(* IEC 61131-3 sources: plcassist-cli/packages/volt-lsp-iec/test-corpus/lenze-mid/Device/Plc Logic/Application/Library Manager/L_MC1P_MotionControlBasic (part 8) *)

(* ---- MC_READBOOLPARAMETER.fb ---- *)
FUNCTION_BLOCK MC_READBOOLPARAMETER EXTENDS L_MC1P_Template_NoAxis
VAR_INPUT
	AXIS : L_MC1P_IMCParameterAccess;
	ENABLE : BOOL;
	PARAMETERNUMBER : DINT;
END_VAR
VAR_OUTPUT
	VALID : BOOL;
	BUSY : BOOL;
	ERROR : BOOL;
	ERRORID : L_IE1P_Error;
	VALUE : BOOL;
END_VAR
VAR
	XENABLEOLD : BOOL := FALSE;
	PARAMETERNUMBEROLD : DINT := 0;
	L_DCO_READDRIVEPARAMETER1 : L_DCO_ReadDriveParameter;
	TIMERREADCYCLE : TON;
	TCYCLETIME : TIME := TIME#1ms;
	XERRORHOLD : BOOL;
	EERRORIDHOLD : L_IE1P_Error;
	PAXISREF : POINTER TO AXIS_REF;
	PINSTANCE : POINTER TO BYTE;
	EAXISTYPE : L_MC1P_AxisType;
	AXISOLD : L_MC1P_IMCParameterAccess;
	_MCCALL : L_UM1P_MCMultipleCall;
	INPUTDATA : ARRAY [1.._MCCall.c_BufferDepthInput] OF L_MC1P_ReadBoolParameterInput;
	OUTPUTDATA : ARRAY [1.._MCCall.c_BufferDepthOutput] OF L_MC1P_ReadBoolParameterOutput;
	POUTPUTDATA : POINTER TO L_MC1P_ReadBoolParameterOutput;
	XAXISTASKIDXVALID : BOOL;
	ITFSETPOINTINFO : L_UM1P_ISetpointInfo;
	IAXISTASKIDX : INT;
	READCYCLE : TIME;
END_VAR
END_FUNCTION_BLOCK

METHOD FB_RESET : BOOL
END_METHOD

METHOD CALLFUNCTION
VAR_INPUT
	UIINPUTDATAIDX : UINT;
	UIOUTPUTDATAIDX : UINT;
END_VAR
END_METHOD

METHOD COPYINPUTS : BOOL
VAR_INPUT
	IDX : WORD;
END_VAR
END_METHOD

METHOD COPYOUTPUTS : BOOL
VAR_INPUT
	IDX : WORD;
END_VAR
END_METHOD

METHOD FUNCTIONWASCALLEDTWICE : BOOL
VAR_INPUT
	IDX : WORD;
END_VAR
END_METHOD

METHOD HANDLESTANDARDCALL : BOOL
END_METHOD

METHOD SYNCOUTPUTS
VAR_INPUT
	UICOPYOUTPUTFROMIDX : UINT;
	UICOPYOUTPUTTOIDX : UINT;
END_VAR
END_METHOD

(* ---- MC_READMOTIONSTATE.fb ---- *)
FUNCTION_BLOCK MC_READMOTIONSTATE EXTENDS L_MC1P_Template
VAR_INPUT
	ENABLE : BOOL;
	SOURCE : MC_SOURCE;
END_VAR
VAR_OUTPUT
	VALID : BOOL;
	BUSY : BOOL;
	ERROR : BOOL;
	ERRORID : L_IE1P_Error;
	CONSTANTVELOCITY : BOOL;
	ACCELERATING : BOOL;
	DECELERATING : BOOL;
	DIRECTIONPOSITIVE : BOOL;
	DIRECTIONNEGATIVE : BOOL;
	INPOSITION : BOOL;
	STANDSTILLSETVELOCITY : BOOL;
	STANDSTILLACTVELOCITY : BOOL;
END_VAR
VAR
	READ : L_MC1P_ReadMotionState_Internal;
	_MCCALL : L_UM1P_MCMultipleCall;
	INPUTDATA : ARRAY [1.._MCCall.c_BufferDepthInput] OF L_MC1P_ReadMotionStateInput;
	OUTPUTDATA : ARRAY [1.._MCCall.c_BufferDepthOutput] OF L_MC1P_ReadMotionStateOutput;
END_VAR
END_FUNCTION_BLOCK

METHOD CALLFUNCTION
VAR_INPUT
	UIINPUTDATAIDX : UINT;
	UIOUTPUTDATAIDX : UINT;
END_VAR
END_METHOD

METHOD COPYINPUTS : BOOL
VAR_INPUT
	IDX : WORD;
END_VAR
END_METHOD

METHOD COPYOUTPUTS : BOOL
VAR_INPUT
	IDX : WORD;
END_VAR
END_METHOD

METHOD FUNCTIONWASCALLEDTWICE : BOOL
VAR_INPUT
	IDX : WORD;
END_VAR
END_METHOD

METHOD HANDLESTANDARDCALL : BOOL
END_METHOD

METHOD SYNCOUTPUTS
VAR_INPUT
	UICOPYOUTPUTFROMIDX : UINT;
	UICOPYOUTPUTTOIDX : UINT;
END_VAR
END_METHOD

(* ---- MC_READPARAMETER.fb ---- *)
FUNCTION_BLOCK MC_READPARAMETER EXTENDS L_MC1P_Template_NoAxis
VAR_INPUT
	AXIS : L_MC1P_IMCParameterAccess;
	ENABLE : BOOL;
	PARAMETERNUMBER : DINT;
END_VAR
VAR_OUTPUT
	VALID : BOOL;
	BUSY : BOOL;
	ERROR : BOOL;
	ERRORID : L_IE1P_Error;
	VALUE : LREAL;
END_VAR
VAR
	READ : L_MC1P_ReadParameter_Internal;
	TCYCLETIME : TIME := TIME#1ms;
	_MCCALL : L_UM1P_MCMultipleCall;
	INPUTDATA : ARRAY [1.._MCCall.c_BufferDepthInput] OF L_MC1P_ReadParameterInput;
	OUTPUTDATA : ARRAY [1.._MCCall.c_BufferDepthOutput] OF L_MC1P_ReadParameterOutput;
	PINPUTDATA : POINTER TO L_MC1P_ReadParameterInput;
	ITFSETPOINTINFO : L_UM1P_ISetpointInfo;
	XAXISTASKIDXVALID : BOOL;
	IAXISTASKIDX : INT;
	READCYCLE : TIME;
END_VAR
END_FUNCTION_BLOCK

METHOD CALLFUNCTION
VAR_INPUT
	UIINPUTDATAIDX : UINT;
	UIOUTPUTDATAIDX : UINT;
END_VAR
END_METHOD

METHOD COPYINPUTS : BOOL
VAR_INPUT
	IDX : WORD;
END_VAR
END_METHOD

METHOD COPYOUTPUTS : BOOL
VAR_INPUT
	IDX : WORD;
END_VAR
END_METHOD

METHOD FUNCTIONWASCALLEDTWICE : BOOL
VAR_INPUT
	IDX : WORD;
END_VAR
END_METHOD

METHOD HANDLESTANDARDCALL : BOOL
END_METHOD

METHOD SYNCOUTPUTS
VAR_INPUT
	UICOPYOUTPUTFROMIDX : UINT;
	UICOPYOUTPUTTOIDX : UINT;
END_VAR
END_METHOD

(* ---- MC_READSTATUS.fb ---- *)
FUNCTION_BLOCK MC_READSTATUS EXTENDS L_MC1P_Template
VAR_INPUT
	ENABLE : BOOL;
END_VAR
VAR_OUTPUT
	VALID : BOOL;
	BUSY : BOOL;
	ERROR : BOOL;
	ERRORID : L_IE1P_Error;
	ERRORSTOP : BOOL;
	DISABLED : BOOL;
	STOPPING : BOOL;
	HOMING : BOOL;
	STANDSTILL : BOOL;
	DISCRETEMOTION : BOOL;
	CONTINUOUSMOTION : BOOL;
	SYNCHRONIZEDMOTION : BOOL;
	CONSTANTVELOCITY : BOOL;
	ACCELERATING : BOOL;
	DECELERATING : BOOL;
	INPOSITION : BOOL;
END_VAR
VAR
	XENABLEOLD : BOOL := FALSE;
	_MCCALL : L_UM1P_MCMultipleCall;
	INPUTDATA : ARRAY [1.._MCCall.c_BufferDepthInput] OF L_MC1P_ReadStatusInput;
	OUTPUTDATA : ARRAY [1.._MCCall.c_BufferDepthOutput] OF L_MC1P_ReadStatusOutput;
	POUTPUTDATA : POINTER TO L_MC1P_ReadStatusOutput;
END_VAR
END_FUNCTION_BLOCK

METHOD FB_RESET : BOOL
END_METHOD

METHOD CALLFUNCTION
VAR_INPUT
	UIINPUTDATAIDX : UINT;
	UIOUTPUTDATAIDX : UINT;
END_VAR
END_METHOD

METHOD COPYINPUTS : BOOL
VAR_INPUT
	IDX : WORD;
END_VAR
END_METHOD

METHOD COPYOUTPUTS : BOOL
VAR_INPUT
	IDX : WORD;
END_VAR
END_METHOD

METHOD FUNCTIONWASCALLEDTWICE : BOOL
VAR_INPUT
	IDX : WORD;
END_VAR
END_METHOD

METHOD HANDLESTANDARDCALL : BOOL
END_METHOD

METHOD SYNCOUTPUTS
VAR_INPUT
	UICOPYOUTPUTFROMIDX : UINT;
	UICOPYOUTPUTTOIDX : UINT;
END_VAR
END_METHOD

(* ---- MC_RESET.fb ---- *)
FUNCTION_BLOCK MC_RESET EXTENDS L_MC1P_Template
VAR_INPUT
	EXECUTE : BOOL;
END_VAR
VAR_OUTPUT
	DONE : BOOL;
	BUSY : BOOL;
	ERROR : BOOL;
	ERRORID : L_IE1P_Error;
END_VAR
VAR
	RESET : L_MC1P_Reset_Internal;
	RESETINPUT : L_MC1P_ResetInput;
	RESETOUTPUT : L_MC1P_ResetOutput;
	_MCCALL : L_UM1P_MCMultipleCall := STRUCT(itfMCCall := THIS^);
	INPUTDATA : ARRAY [1.._MCCall.c_BufferDepthInput] OF L_MC1P_ResetInput;
	OUTPUTDATA : ARRAY [1.._MCCall.c_BufferDepthOutput] OF L_MC1P_ResetOutput;
	POUTPUTDATA : POINTER TO L_MC1P_ResetOutput;
END_VAR
END_FUNCTION_BLOCK

METHOD CALLFUNCTION
VAR_INPUT
	UIINPUTDATAIDX : UINT;
	UIOUTPUTDATAIDX : UINT;
END_VAR
END_METHOD

METHOD COPYINPUTS : BOOL
VAR_INPUT
	IDX : WORD;
END_VAR
END_METHOD

METHOD COPYOUTPUTS : BOOL
VAR_INPUT
	IDX : WORD;
END_VAR
END_METHOD

METHOD FUNCTIONWASCALLEDTWICE : BOOL
VAR_INPUT
	IDX : WORD;
END_VAR
END_METHOD

METHOD HANDLESTANDARDCALL : BOOL
END_METHOD

METHOD SYNCOUTPUTS
VAR_INPUT
	UICOPYOUTPUTFROMIDX : UINT;
	UICOPYOUTPUTTOIDX : UINT;
END_VAR
END_METHOD

(* ---- MC_SETOVERRIDE.fb ---- *)
FUNCTION_BLOCK MC_SETOVERRIDE EXTENDS L_MC1P_Template
VAR_INPUT
	ENABLE : BOOL;
	VELFACTOR : LREAL := 1.0;
	ACCFACTOR : LREAL := 1.0;
	JERKFACTOR : LREAL := 1.0;
END_VAR
VAR_OUTPUT
	ENABLED : BOOL;
	BUSY : BOOL;
	ERROR : BOOL;
	ERRORID : L_IE1P_Error;
END_VAR
VAR
	OVERRIDE : L_MC1P_SetOverride_Internal;
	_MCCALL : L_UM1P_MCMultipleCall;
	INPUTDATA : ARRAY [1.._MCCall.c_BufferDepthInput] OF L_MC1P_SetOverrideInput;
	OUTPUTDATA : ARRAY [1.._MCCall.c_BufferDepthOutput] OF L_MC1P_SetOverrideOutput;
END_VAR
END_FUNCTION_BLOCK

METHOD CALLFUNCTION
VAR_INPUT
	UIINPUTDATAIDX : UINT;
	UIOUTPUTDATAIDX : UINT;
END_VAR
END_METHOD

METHOD COPYINPUTS : BOOL
VAR_INPUT
	IDX : WORD;
END_VAR
END_METHOD

METHOD COPYOUTPUTS : BOOL
VAR_INPUT
	IDX : WORD;
END_VAR
END_METHOD

METHOD FUNCTIONWASCALLEDTWICE : BOOL
VAR_INPUT
	IDX : WORD;
END_VAR
END_METHOD

METHOD HANDLESTANDARDCALL : BOOL
END_METHOD

METHOD SYNCOUTPUTS
VAR_INPUT
	UICOPYOUTPUTFROMIDX : UINT;
	UICOPYOUTPUTTOIDX : UINT;
END_VAR
END_METHOD

(* ---- MC_SETPOSITION.fb ---- *)
FUNCTION_BLOCK MC_SETPOSITION EXTENDS L_MC1P_Template
VAR_INPUT
	EXECUTE : BOOL;
	POSITION : LREAL;
	RELATIVE : BOOL;
	EXECUTIONMODE : MC_EXECUTION_MODE := MC_EXECUTION_MODE.mcImmediately;
	RESTARTPOSITIONING : BOOL := FALSE;
	USESETTINGSFROMHOMINGMODE : BOOL := FALSE;
END_VAR
VAR_OUTPUT
	DONE : BOOL;
	BUSY : BOOL;
	ERROR : BOOL;
	ERRORID : L_IE1P_Error;
END_VAR
VAR
	XEXECUTEOLD : BOOL;
	XCALLFROMAXESGROUP : BOOL;
	LRDUMMY : LREAL;
	XDISABLELOGMESSAGE : BOOL := FALSE;
	_MCCALL : L_UM1P_MCMultipleCall;
	INPUTDATA : ARRAY [1.._MCCall.c_BufferDepthInput] OF L_MC1P_SetPositionInput;
	OUTPUTDATA : ARRAY [1.._MCCall.c_BufferDepthOutput] OF L_MC1P_SetPositionOutput;
	DISABLELOGMESSAGE : BOOL;
END_VAR
END_FUNCTION_BLOCK

METHOD SETCALLFROMAXESGROUP
VAR_INPUT
	XSETCALLFROMAXESGROUP : BOOL;
END_VAR
END_METHOD

METHOD CALLFUNCTION
VAR_INPUT
	UIINPUTDATAIDX : UINT;
	UIOUTPUTDATAIDX : UINT;
END_VAR
END_METHOD

METHOD COPYINPUTS : BOOL
VAR_INPUT
	IDX : WORD;
END_VAR
END_METHOD

METHOD COPYOUTPUTS : BOOL
VAR_INPUT
	IDX : WORD;
END_VAR
END_METHOD

METHOD FUNCTIONWASCALLEDTWICE : BOOL
VAR_INPUT
	IDX : WORD;
END_VAR
END_METHOD

METHOD HANDLESTANDARDCALL : BOOL
END_METHOD

METHOD SYNCOUTPUTS
VAR_INPUT
	UICOPYOUTPUTFROMIDX : UINT;
	UICOPYOUTPUTTOIDX : UINT;
END_VAR
END_METHOD

(* ---- MC_STOP.fb ---- *)
FUNCTION_BLOCK MC_STOP EXTENDS L_MC1P_Template_Licence_150
VAR_INPUT
	EXECUTE : BOOL;
	DECELERATION : LREAL;
	JERK : LREAL;
END_VAR
VAR_OUTPUT
	DONE : BOOL;
	BUSY : BOOL;
	COMMANDABORTED : BOOL;
	ERROR : BOOL;
	ERRORID : L_IE1P_Error;
END_VAR
VAR
	STOP : L_MC1P_Stop_Internal;
	_MCCALL : L_UM1P_MCMultipleCall;
	INPUTDATA : ARRAY [1.._MCCall.c_BufferDepthInput] OF L_MC1P_StopInput;
	OUTPUTDATA : ARRAY [1.._MCCall.c_BufferDepthOutput] OF L_MC1P_StopOutput;
	PROFILETIME : TIME;
	REMAININGTIMEOFPROFILE : LREAL;
	REMAININGTIMEOFPROFILEAVAILABLE : BOOL;
END_VAR
END_FUNCTION_BLOCK

METHOD CALLFUNCTION
VAR_INPUT
	UIINPUTDATAIDX : UINT;
	UIOUTPUTDATAIDX : UINT;
END_VAR
END_METHOD

METHOD COPYINPUTS : BOOL
VAR_INPUT
	IDX : WORD;
END_VAR
END_METHOD

METHOD COPYOUTPUTS : BOOL
VAR_INPUT
	IDX : WORD;
END_VAR
END_METHOD

METHOD FUNCTIONWASCALLEDTWICE : BOOL
VAR_INPUT
	IDX : WORD;
END_VAR
END_METHOD

METHOD HANDLESTANDARDCALL : BOOL
END_METHOD

METHOD SYNCOUTPUTS
VAR_INPUT
	UICOPYOUTPUTFROMIDX : UINT;
	UICOPYOUTPUTTOIDX : UINT;
END_VAR
END_METHOD

(* ---- MC_TOUCHPROBE.fb ---- *)
FUNCTION_BLOCK MC_TOUCHPROBE EXTENDS L_MC1P_Template
VAR_INPUT
	EXECUTE : BOOL;
	WINDOWONLY : BOOL;
	FIRSTPOSITION : LREAL;
	LASTPOSITION : LREAL;
END_VAR
VAR_OUTPUT
	DONE : BOOL;
	BUSY : BOOL;
	COMMANDABORTED : BOOL;
	ERROR : BOOL;
	ERRORID : L_IE1P_Error;
	ACTIVATIONLEVEL : BOOL;
	ACTIVATIONLEVELVALID : BOOL;
	VALUESTORED_POSEDGE : BOOL;
	RECPOSITION_POSEDGE : LREAL;
	VALUESTORED_NEGEDGE : BOOL;
	RECPOSITION_NEGEDGE : LREAL;
	NEWVALUESTORED_POSEDGE : BOOL;
	NEWVALUESTORED_NEGEDGE : BOOL;
	RECDATA : L_MC1P_TpReceiveData;
END_VAR
VAR_IN_OUT
	TRIGGERINPUT : MC_TRIGGER_REF;
END_VAR
VAR
	TP : L_MC1P_TouchProbe_Internal;
	_MCCALL : L_UM1P_MCMultipleCall := STRUCT(itfMCCall := THIS^);
	INPUTDATA : ARRAY [1.._MCCall.c_BufferDepthInput] OF L_MC1P_TouchProbeInput;
	OUTPUTDATA : ARRAY [1.._MCCall.c_BufferDepthOutput] OF L_MC1P_TouchProbeOutput;
	_FB_SEMA : L_MC1P_CriticalSection;
	_DWUPDATETIME : DWORD;
	DWACTTIMESTAMPSAVE : DWORD;
	XMULTICOREOPTION : BOOL;
END_VAR
END_FUNCTION_BLOCK

METHOD GETACTTPRECEIVEDATA : L_MC1P_TpReceiveData
END_METHOD

METHOD ISUPTODATE : BOOL
VAR_INPUT
	DWUPDATETIME : DWORD;
END_VAR
END_METHOD

METHOD RECDATAISVALID : BOOL
VAR_IN_OUT
	SCRECDATA : L_MC1P_TpReceiveData;
END_VAR
END_METHOD

METHOD REQUESTINTERFACE : BOOL
VAR_INPUT
	ID : DINT;
	PITFUNKNOWN : POINTER TO L_UBUP_IUnknown;
END_VAR
END_METHOD

METHOD CALLFUNCTION
VAR_INPUT
	UIINPUTDATAIDX : UINT;
	UIOUTPUTDATAIDX : UINT;
END_VAR
END_METHOD

METHOD COPYINPUTS : BOOL
VAR_INPUT
	IDX : WORD;
END_VAR
END_METHOD

METHOD COPYOUTPUTS : BOOL
VAR_INPUT
	IDX : WORD;
END_VAR
END_METHOD

METHOD FUNCTIONWASCALLEDTWICE : BOOL
VAR_INPUT
	IDX : WORD;
END_VAR
END_METHOD

METHOD HANDLESTANDARDCALL : BOOL
END_METHOD

METHOD SYNCOUTPUTS
VAR_INPUT
	UICOPYOUTPUTFROMIDX : UINT;
	UICOPYOUTPUTTOIDX : UINT;
END_VAR
END_METHOD

(* ---- MC_WRITEBOOLPARAMETER.fb ---- *)
FUNCTION_BLOCK MC_WRITEBOOLPARAMETER EXTENDS L_MC1P_Template_NoAxis
VAR_INPUT
	AXIS : L_MC1P_IMCParameterAccess;
	EXECUTE : BOOL;
	PARAMETERNUMBER : DINT;
	VALUE : BOOL;
	EXECUTIONMODE : MC_EXECUTION_MODE;
END_VAR
VAR_OUTPUT
	DONE : BOOL;
	BUSY : BOOL;
	ERROR : BOOL;
	ERRORID : L_IE1P_Error;
END_VAR
VAR
	XEXECUTEOLD : BOOL := FALSE;
	XRESETOUTPUT : BOOL := FALSE;
	L_DCO_WRITEDRIVEPARAMETER1 : L_DCO_WriteDriveParameter;
	WERRORID_INT : WORD;
	AXISOLD : L_MC1P_IMCParameterAccess;
	PAXISREF : POINTER TO AXIS_REF;
	XWRITEPARAMETER : BOOL;
	PINSTANCE : POINTER TO BYTE;
	EAXISTYPE : L_MC1P_AxisType;
	_MCCALL : L_UM1P_MCMultipleCall;
	INPUTDATA : ARRAY [1.._MCCall.c_BufferDepthInput] OF L_MC1P_WriteBoolParameterInput;
	OUTPUTDATA : ARRAY [1.._MCCall.c_BufferDepthOutput] OF L_MC1P_WriteBoolParameterOutput;
	POUTPUTDATA : POINTER TO L_MC1P_WriteBoolParameterOutput;
	ITFSETPOINTINFO : L_UM1P_ISetpointInfo;
	XAXISTASKIDXVALID : BOOL;
	IAXISTASKIDX : INT;
END_VAR
END_FUNCTION_BLOCK

METHOD FB_RESET : BOOL
END_METHOD

METHOD CALLFUNCTION
VAR_INPUT
	UIINPUTDATAIDX : UINT;
	UIOUTPUTDATAIDX : UINT;
END_VAR
END_METHOD

METHOD COPYINPUTS : BOOL
VAR_INPUT
	IDX : WORD;
END_VAR
END_METHOD

METHOD COPYOUTPUTS : BOOL
VAR_INPUT
	IDX : WORD;
END_VAR
END_METHOD

METHOD FUNCTIONWASCALLEDTWICE : BOOL
VAR_INPUT
	IDX : WORD;
END_VAR
END_METHOD

METHOD HANDLESTANDARDCALL : BOOL
END_METHOD

METHOD SYNCOUTPUTS
VAR_INPUT
	UICOPYOUTPUTFROMIDX : UINT;
	UICOPYOUTPUTTOIDX : UINT;
END_VAR
END_METHOD

(* ---- MC_WRITEPARAMETER.fb ---- *)
FUNCTION_BLOCK MC_WRITEPARAMETER EXTENDS L_MC1P_Template_NoAxis
VAR_INPUT
	AXIS : L_MC1P_IMCParameterAccess;
	EXECUTE : BOOL;
	PARAMETERNUMBER : DINT;
	VALUE : LREAL;
	EXECUTIONMODE : MC_EXECUTION_MODE;
END_VAR
VAR_OUTPUT
	DONE : BOOL;
	BUSY : BOOL;
	ERROR : BOOL;
	ERRORID : L_IE1P_Error;
END_VAR
VAR
	XEXECUTEOLD : BOOL := FALSE;
	XRESETOUTPUT : BOOL := FALSE;
	AXISOLD : L_MC1P_IMCParameterAccess;
	L_DCO_WRITEDRIVEPARAMETER1 : L_DCO_WriteDriveParameter;
	DWPARAMETERNUMBERINT : DWORD;
	WERRORID_INT : WORD;
	PAXISREF : POINTER TO AXIS_REF;
	PINSTANCE : POINTER TO BYTE;
	EAXISTYPE : L_MC1P_AxisType;
	_MCCALL : L_UM1P_MCMultipleCall;
	INPUTDATA : ARRAY [1.._MCCall.c_BufferDepthInput] OF L_MC1P_WriteParameterInput;
	OUTPUTDATA : ARRAY [1.._MCCall.c_BufferDepthOutput] OF L_MC1P_WriteParameterOutput;
	POUTPUTDATA : POINTER TO L_MC1P_WriteParameterOutput;
	ITFSETPOINTINFO : L_UM1P_ISetpointInfo;
	XAXISTASKIDXVALID : BOOL;
	IAXISTASKIDX : INT;
END_VAR
END_FUNCTION_BLOCK

METHOD FB_RESET : BOOL
END_METHOD

METHOD CALLFUNCTION
VAR_INPUT
	UIINPUTDATAIDX : UINT;
	UIOUTPUTDATAIDX : UINT;
END_VAR
END_METHOD

METHOD COPYINPUTS : BOOL
VAR_INPUT
	IDX : WORD;
END_VAR
END_METHOD

METHOD COPYOUTPUTS : BOOL
VAR_INPUT
	IDX : WORD;
END_VAR
END_METHOD

METHOD FUNCTIONWASCALLEDTWICE : BOOL
VAR_INPUT
	IDX : WORD;
END_VAR
END_METHOD

METHOD HANDLESTANDARDCALL : BOOL
END_METHOD

METHOD SYNCOUTPUTS
VAR_INPUT
	UICOPYOUTPUTFROMIDX : UINT;
	UICOPYOUTPUTTOIDX : UINT;
END_VAR
END_METHOD

(* ---- TEXTLIST.fb ---- *)
FUNCTION_BLOCK TEXTLIST
VAR
	M_TEXTLISTFILE : STRING(255);
	_STNAMESPACE : STRING;
END_VAR
END_FUNCTION_BLOCK
